(* Schneider Machine Expert - Basic project New project, file version 2.9.0.0 *)
(* ProjectInformations: Name=New project *)

HARDWARE
  Cpu 0: TM221M16R/G
  ModuleExtensionObject 0: TM3DI16K
  ModuleExtensionObject 1: TM3DQ16R/G
  EthernetConfiguration: NetworkName=M221, IpAllocationMode=FixedAddress, IpAddress=0.0.0.0, SubnetMask=0.0.0.0
  SerialLineConfiguration: Baud=Baud19200, Parity=ParityEven, DataBits=DataBits8, StopBits=StopBits1, PhysicalMedium=PhysicalMediumRs485, TransmissionMode=TransmissionModeModbusRtu, SlaveId=1, Addressing=SlaveAddressing
  MastTask: UsePeriodScanMode=false, PeriodScan=100
  FastTask: Period=255
  CpuBehavior: StartingMode=StartAsPreviousState, AutoSaveRamOnEeprom=true, WatchdogPeriod=250

SYMBOLS  (address, symbol, comment, settings)
  %M0       C_1
  %M1       C_2
  %M2       DM_PMP_STAT
  %I0.0     A
  %I0.1     B
  %I0.2     DI_PMP_START
  %I0.3     DI_PMP_STOP
  %Q2.0     C
  %Q2.1     DQ_PMP_RUN

POU New POU
  (* SectionNumber=1 *)

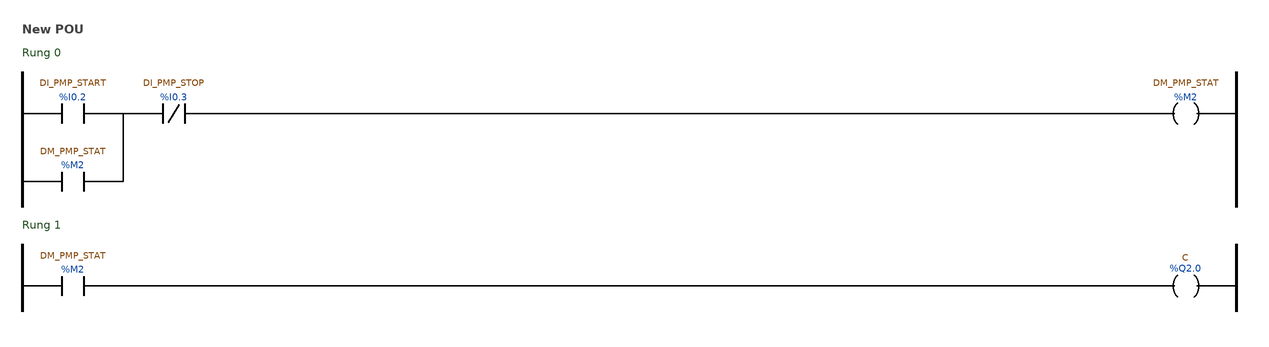

// Rung 0
  LD %I0.2                (* DI_PMP_START *)
  OR %M2                  (* DM_PMP_STAT *)
  ANDN %I0.3              (* DI_PMP_STOP *)
  ST %M2                  (* DM_PMP_STAT *)
  // as ST:
  //   DM_PMP_STAT := (DI_PMP_START OR DM_PMP_STAT) AND NOT DI_PMP_STOP;

// Rung 1
  LD %M2                  (* DM_PMP_STAT *)
  ST %Q2.0                (* C *)
  // as ST:
  //   C := DM_PMP_STAT;
